(* Logix 5000 project; controller CIP vendor 1 type 14 code 106 rev 20.12; software revision 20.06; part 10 of 13 *)
(* tags used below, declared in another part *)
   MOA_OFF : DINT[10];
   MOA_ON : DINT[10];
   PV_Output_Status : INT[10];
   PV_Output_Status_IND : INT[10,16];
   PV_Status_Bit : BOOL;
   PV_Valve_Input_Status_IND : INT[10,16];
(* MainProgram, continued *)

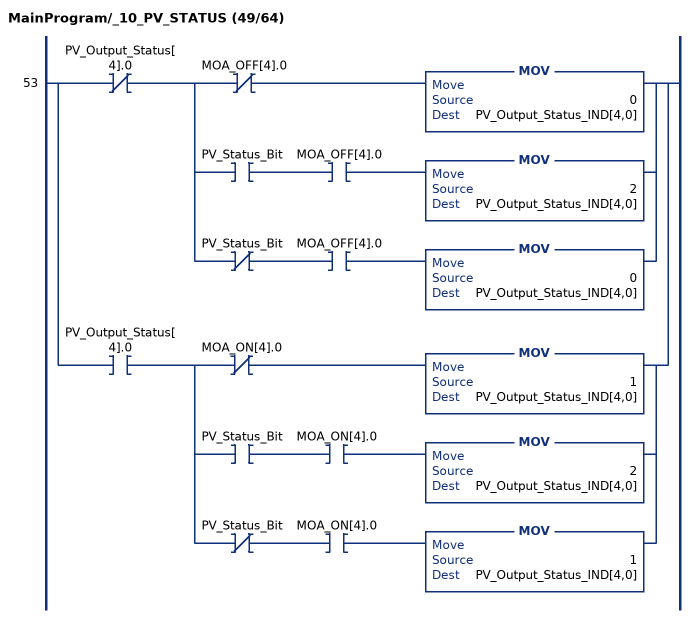
   [picture p181: MainProgram/_10_PV_STATUS rungs 53-53]
   53: [XIO(PV_Output_Status[4].0) [XIO(MOA_OFF[4].0) MOV(0,PV_Output_Status_IND[4,0]) ,XIC(PV_Status_Bit) XIC(MOA_OFF[4].0) MOV(2,PV_Output_Status_IND[4,0]) ,XIO(PV_Status_Bit) XIC(MOA_OFF[4].0) MOV(0,PV_Output_Status_IND[4,0]) ] ,XIC(PV_Output_Status[4].0) [XIO(MOA_ON[4].0) MOV(1,PV_Output_Status_IND[4,0]) ,XIC(PV_Status_Bit) XIC(MOA_ON[4].0) MOV(2,PV_Output_Status_IND[4,0]) ,XIO(PV_Status_Bit) XIC(MOA_ON[4].0) MOV(1,PV_Output_Status_IND[4,0]) ] ];
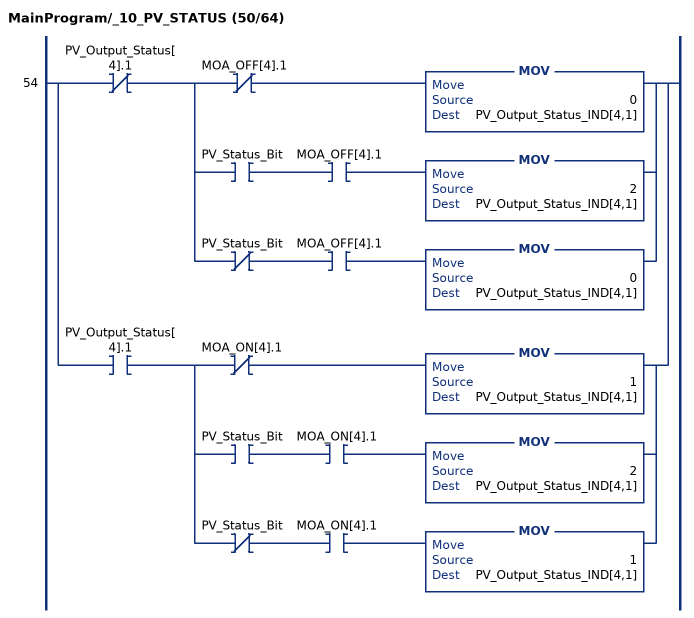
   54: [XIO(PV_Output_Status[4].1) [XIO(MOA_OFF[4].1) MOV(0,PV_Output_Status_IND[4,1]) ,XIC(PV_Status_Bit) XIC(MOA_OFF[4].1) MOV(2,PV_Output_Status_IND[4,1]) ,XIO(PV_Status_Bit) XIC(MOA_OFF[4].1) MOV(0,PV_Output_Status_IND[4,1]) ] ,XIC(PV_Output_Status[4].1) [XIO(MOA_ON[4].1) MOV(1,PV_Output_Status_IND[4,1]) ,XIC(PV_Status_Bit) XIC(MOA_ON[4].1) MOV(2,PV_Output_Status_IND[4,1]) ,XIO(PV_Status_Bit) XIC(MOA_ON[4].1) MOV(1,PV_Output_Status_IND[4,1]) ] ];
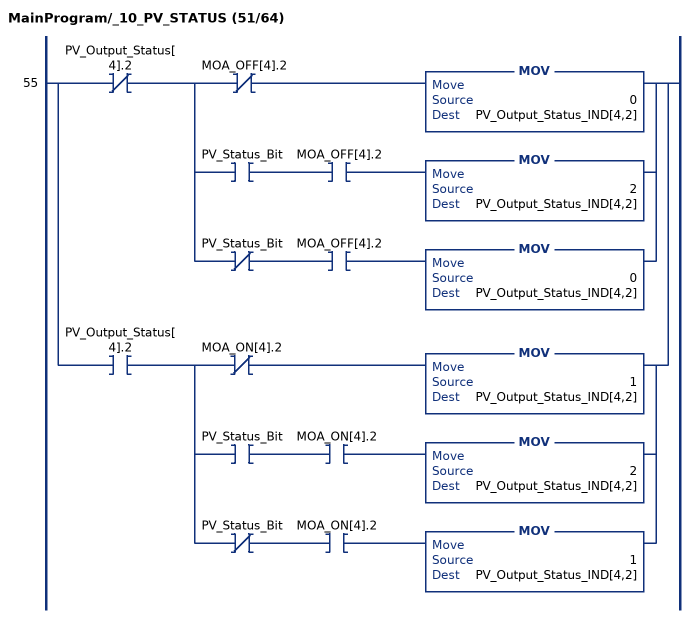
   55: [XIO(PV_Output_Status[4].2) [XIO(MOA_OFF[4].2) MOV(0,PV_Output_Status_IND[4,2]) ,XIC(PV_Status_Bit) XIC(MOA_OFF[4].2) MOV(2,PV_Output_Status_IND[4,2]) ,XIO(PV_Status_Bit) XIC(MOA_OFF[4].2) MOV(0,PV_Output_Status_IND[4,2]) ] ,XIC(PV_Output_Status[4].2) [XIO(MOA_ON[4].2) MOV(1,PV_Output_Status_IND[4,2]) ,XIC(PV_Status_Bit) XIC(MOA_ON[4].2) MOV(2,PV_Output_Status_IND[4,2]) ,XIO(PV_Status_Bit) XIC(MOA_ON[4].2) MOV(1,PV_Output_Status_IND[4,2]) ] ];
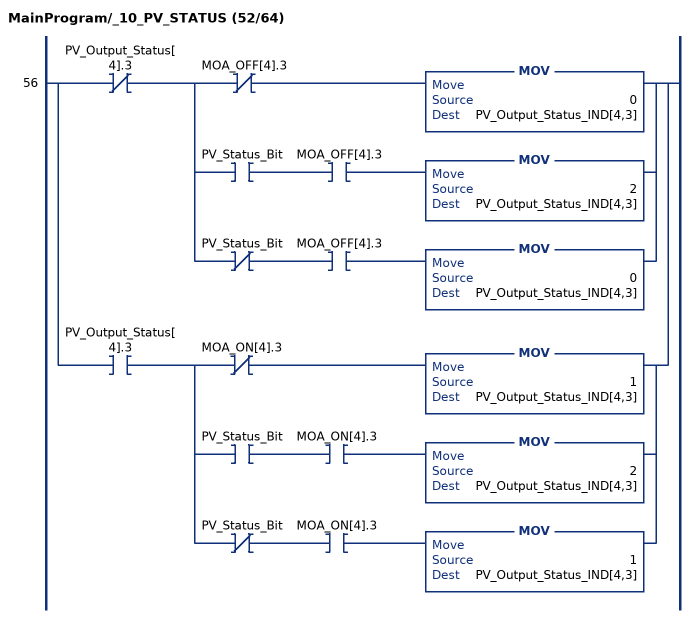
   56: [XIO(PV_Output_Status[4].3) [XIO(MOA_OFF[4].3) MOV(0,PV_Output_Status_IND[4,3]) ,XIC(PV_Status_Bit) XIC(MOA_OFF[4].3) MOV(2,PV_Output_Status_IND[4,3]) ,XIO(PV_Status_Bit) XIC(MOA_OFF[4].3) MOV(0,PV_Output_Status_IND[4,3]) ] ,XIC(PV_Output_Status[4].3) [XIO(MOA_ON[4].3) MOV(1,PV_Output_Status_IND[4,3]) ,XIC(PV_Status_Bit) XIC(MOA_ON[4].3) MOV(2,PV_Output_Status_IND[4,3]) ,XIO(PV_Status_Bit) XIC(MOA_ON[4].3) MOV(1,PV_Output_Status_IND[4,3]) ] ];
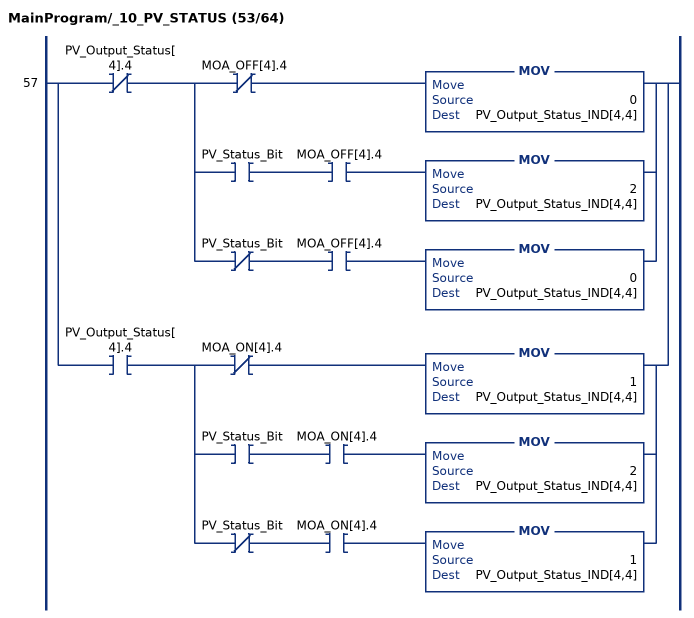
   57: [XIO(PV_Output_Status[4].4) [XIO(MOA_OFF[4].4) MOV(0,PV_Output_Status_IND[4,4]) ,XIC(PV_Status_Bit) XIC(MOA_OFF[4].4) MOV(2,PV_Output_Status_IND[4,4]) ,XIO(PV_Status_Bit) XIC(MOA_OFF[4].4) MOV(0,PV_Output_Status_IND[4,4]) ] ,XIC(PV_Output_Status[4].4) [XIO(MOA_ON[4].4) MOV(1,PV_Output_Status_IND[4,4]) ,XIC(PV_Status_Bit) XIC(MOA_ON[4].4) MOV(2,PV_Output_Status_IND[4,4]) ,XIO(PV_Status_Bit) XIC(MOA_ON[4].4) MOV(1,PV_Output_Status_IND[4,4]) ] ];
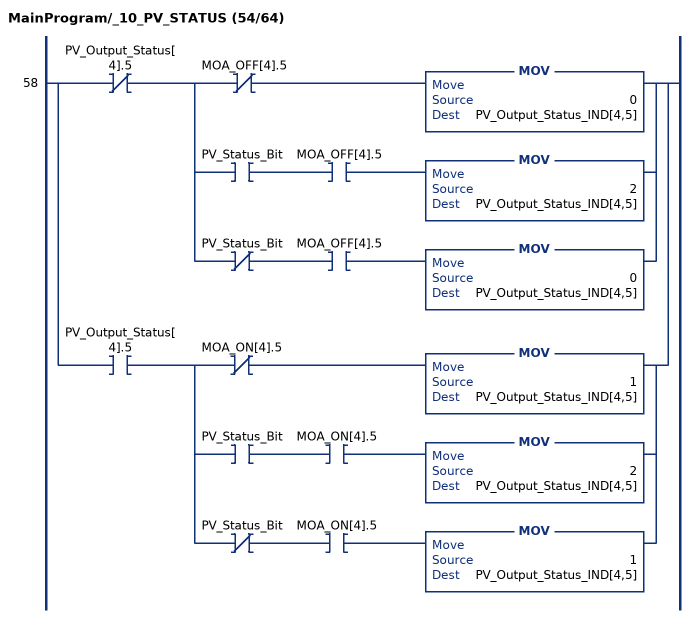
   58: [XIO(PV_Output_Status[4].5) [XIO(MOA_OFF[4].5) MOV(0,PV_Output_Status_IND[4,5]) ,XIC(PV_Status_Bit) XIC(MOA_OFF[4].5) MOV(2,PV_Output_Status_IND[4,5]) ,XIO(PV_Status_Bit) XIC(MOA_OFF[4].5) MOV(0,PV_Output_Status_IND[4,5]) ] ,XIC(PV_Output_Status[4].5) [XIO(MOA_ON[4].5) MOV(1,PV_Output_Status_IND[4,5]) ,XIC(PV_Status_Bit) XIC(MOA_ON[4].5) MOV(2,PV_Output_Status_IND[4,5]) ,XIO(PV_Status_Bit) XIC(MOA_ON[4].5) MOV(1,PV_Output_Status_IND[4,5]) ] ];
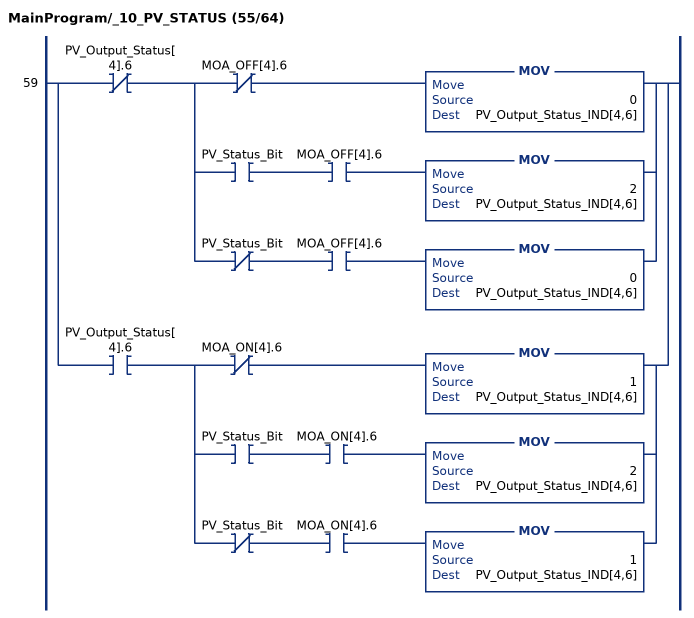
   59: [XIO(PV_Output_Status[4].6) [XIO(MOA_OFF[4].6) MOV(0,PV_Output_Status_IND[4,6]) ,XIC(PV_Status_Bit) XIC(MOA_OFF[4].6) MOV(2,PV_Output_Status_IND[4,6]) ,XIO(PV_Status_Bit) XIC(MOA_OFF[4].6) MOV(0,PV_Output_Status_IND[4,6]) ] ,XIC(PV_Output_Status[4].6) [XIO(MOA_ON[4].6) MOV(1,PV_Output_Status_IND[4,6]) ,XIC(PV_Status_Bit) XIC(MOA_ON[4].6) MOV(2,PV_Output_Status_IND[4,6]) ,XIO(PV_Status_Bit) XIC(MOA_ON[4].6) MOV(1,PV_Output_Status_IND[4,6]) ] ];
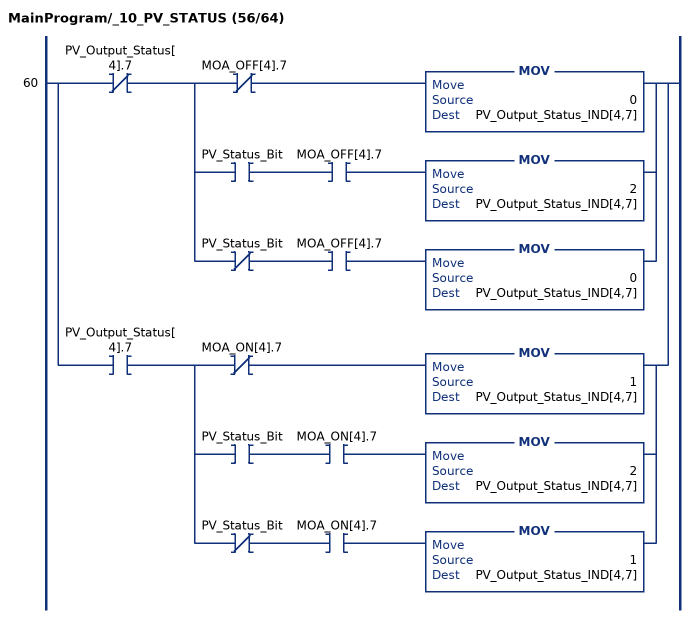
   60: [XIO(PV_Output_Status[4].7) [XIO(MOA_OFF[4].7) MOV(0,PV_Output_Status_IND[4,7]) ,XIC(PV_Status_Bit) XIC(MOA_OFF[4].7) MOV(2,PV_Output_Status_IND[4,7]) ,XIO(PV_Status_Bit) XIC(MOA_OFF[4].7) MOV(0,PV_Output_Status_IND[4,7]) ] ,XIC(PV_Output_Status[4].7) [XIO(MOA_ON[4].7) MOV(1,PV_Output_Status_IND[4,7]) ,XIC(PV_Status_Bit) XIC(MOA_ON[4].7) MOV(2,PV_Output_Status_IND[4,7]) ,XIO(PV_Status_Bit) XIC(MOA_ON[4].7) MOV(1,PV_Output_Status_IND[4,7]) ] ];
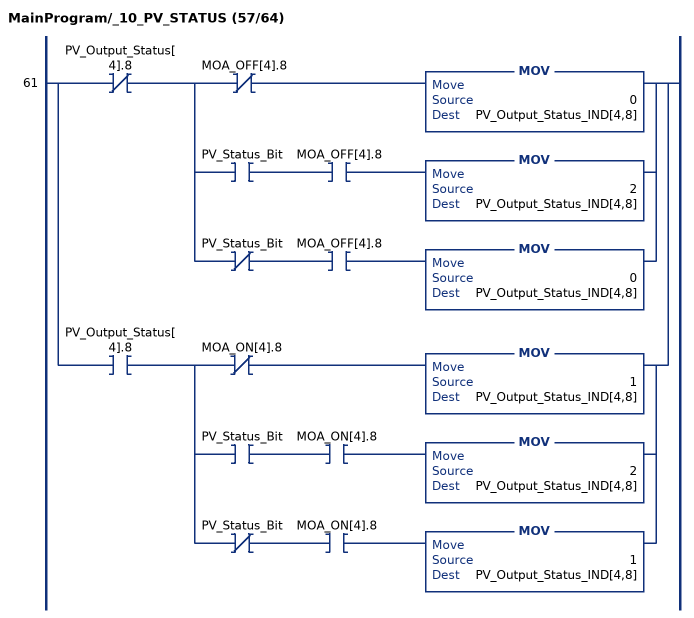
   61: [XIO(PV_Output_Status[4].8) [XIO(MOA_OFF[4].8) MOV(0,PV_Output_Status_IND[4,8]) ,XIC(PV_Status_Bit) XIC(MOA_OFF[4].8) MOV(2,PV_Output_Status_IND[4,8]) ,XIO(PV_Status_Bit) XIC(MOA_OFF[4].8) MOV(0,PV_Output_Status_IND[4,8]) ] ,XIC(PV_Output_Status[4].8) [XIO(MOA_ON[4].8) MOV(1,PV_Output_Status_IND[4,8]) ,XIC(PV_Status_Bit) XIC(MOA_ON[4].8) MOV(2,PV_Output_Status_IND[4,8]) ,XIO(PV_Status_Bit) XIC(MOA_ON[4].8) MOV(1,PV_Output_Status_IND[4,8]) ] ];
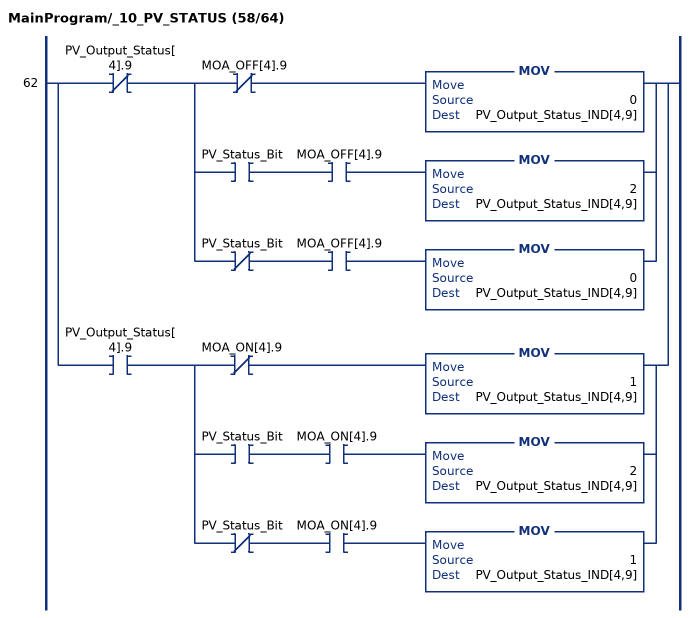
   62: [XIO(PV_Output_Status[4].9) [XIO(MOA_OFF[4].9) MOV(0,PV_Output_Status_IND[4,9]) ,XIC(PV_Status_Bit) XIC(MOA_OFF[4].9) MOV(2,PV_Output_Status_IND[4,9]) ,XIO(PV_Status_Bit) XIC(MOA_OFF[4].9) MOV(0,PV_Output_Status_IND[4,9]) ] ,XIC(PV_Output_Status[4].9) [XIO(MOA_ON[4].9) MOV(1,PV_Output_Status_IND[4,9]) ,XIC(PV_Status_Bit) XIC(MOA_ON[4].9) MOV(2,PV_Output_Status_IND[4,9]) ,XIO(PV_Status_Bit) XIC(MOA_ON[4].9) MOV(1,PV_Output_Status_IND[4,9]) ] ];
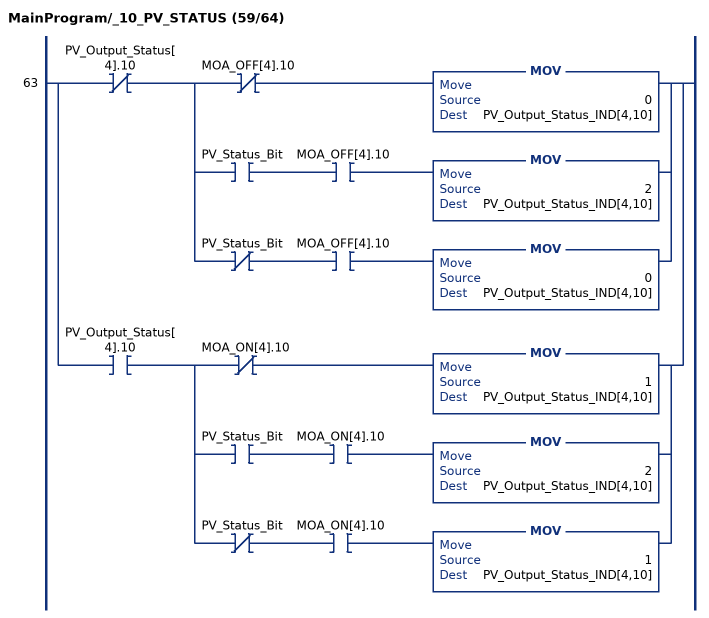
   63: [XIO(PV_Output_Status[4].10) [XIO(MOA_OFF[4].10) MOV(0,PV_Output_Status_IND[4,10]) ,XIC(PV_Status_Bit) XIC(MOA_OFF[4].10) MOV(2,PV_Output_Status_IND[4,10]) ,XIO(PV_Status_Bit) XIC(MOA_OFF[4].10) MOV(0,PV_Output_Status_IND[4,10]) ] ,XIC(PV_Output_Status[4].10) [XIO(MOA_ON[4].10) MOV(1,PV_Output_Status_IND[4,10]) ,XIC(PV_Status_Bit) XIC(MOA_ON[4].10) MOV(2,PV_Output_Status_IND[4,10]) ,XIO(PV_Status_Bit) XIC(MOA_ON[4].10) MOV(1,PV_Output_Status_IND[4,10]) ] ];
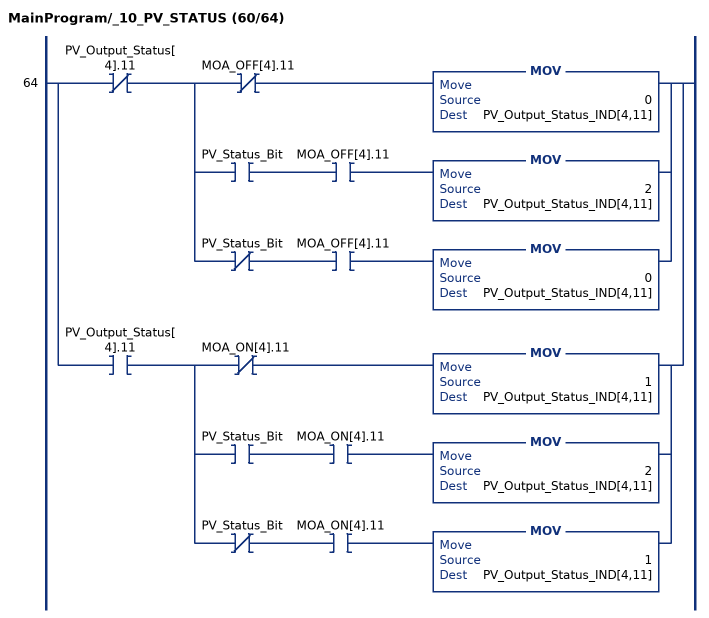
   64: [XIO(PV_Output_Status[4].11) [XIO(MOA_OFF[4].11) MOV(0,PV_Output_Status_IND[4,11]) ,XIC(PV_Status_Bit) XIC(MOA_OFF[4].11) MOV(2,PV_Output_Status_IND[4,11]) ,XIO(PV_Status_Bit) XIC(MOA_OFF[4].11) MOV(0,PV_Output_Status_IND[4,11]) ] ,XIC(PV_Output_Status[4].11) [XIO(MOA_ON[4].11) MOV(1,PV_Output_Status_IND[4,11]) ,XIC(PV_Status_Bit) XIC(MOA_ON[4].11) MOV(2,PV_Output_Status_IND[4,11]) ,XIO(PV_Status_Bit) XIC(MOA_ON[4].11) MOV(1,PV_Output_Status_IND[4,11]) ] ];
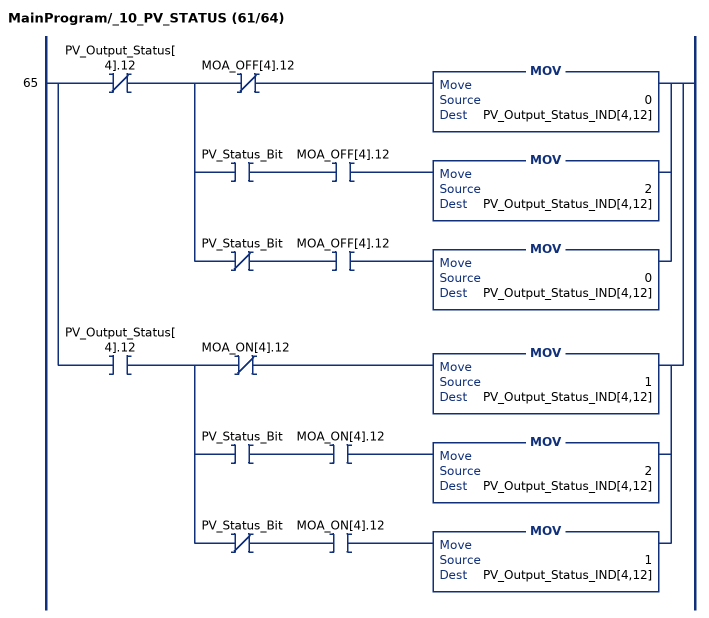
   65: [XIO(PV_Output_Status[4].12) [XIO(MOA_OFF[4].12) MOV(0,PV_Output_Status_IND[4,12]) ,XIC(PV_Status_Bit) XIC(MOA_OFF[4].12) MOV(2,PV_Output_Status_IND[4,12]) ,XIO(PV_Status_Bit) XIC(MOA_OFF[4].12) MOV(0,PV_Output_Status_IND[4,12]) ] ,XIC(PV_Output_Status[4].12) [XIO(MOA_ON[4].12) MOV(1,PV_Output_Status_IND[4,12]) ,XIC(PV_Status_Bit) XIC(MOA_ON[4].12) MOV(2,PV_Output_Status_IND[4,12]) ,XIO(PV_Status_Bit) XIC(MOA_ON[4].12) MOV(1,PV_Output_Status_IND[4,12]) ] ];
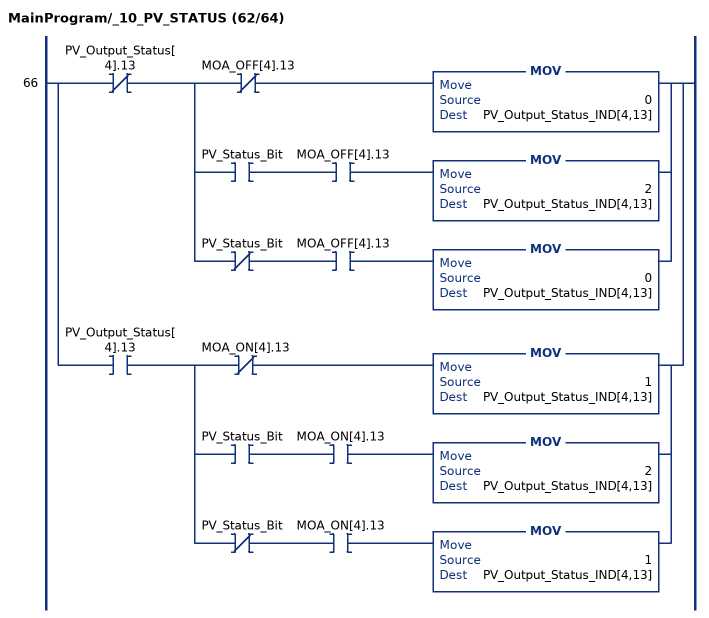
   66: [XIO(PV_Output_Status[4].13) [XIO(MOA_OFF[4].13) MOV(0,PV_Output_Status_IND[4,13]) ,XIC(PV_Status_Bit) XIC(MOA_OFF[4].13) MOV(2,PV_Output_Status_IND[4,13]) ,XIO(PV_Status_Bit) XIC(MOA_OFF[4].13) MOV(0,PV_Output_Status_IND[4,13]) ] ,XIC(PV_Output_Status[4].13) [XIO(MOA_ON[4].13) MOV(1,PV_Output_Status_IND[4,13]) ,XIC(PV_Status_Bit) XIC(MOA_ON[4].13) MOV(2,PV_Output_Status_IND[4,13]) ,XIO(PV_Status_Bit) XIC(MOA_ON[4].13) MOV(1,PV_Output_Status_IND[4,13]) ] ];
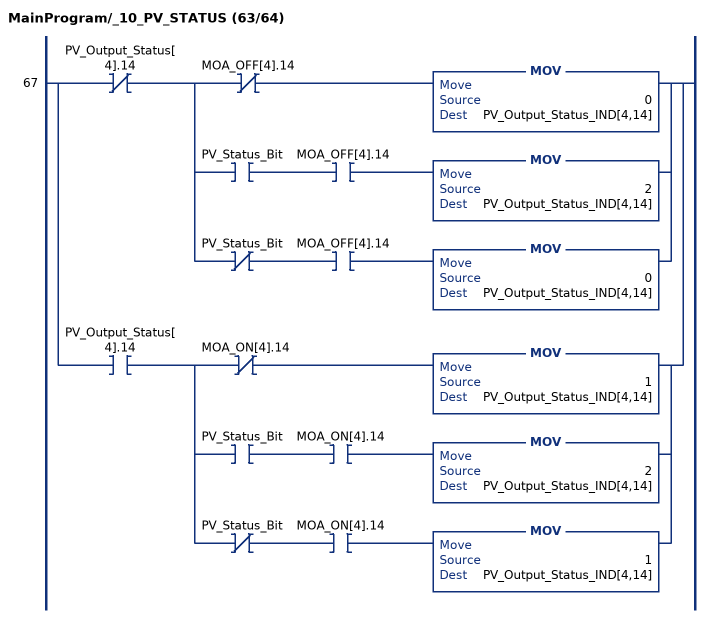
   67: [XIO(PV_Output_Status[4].14) [XIO(MOA_OFF[4].14) MOV(0,PV_Output_Status_IND[4,14]) ,XIC(PV_Status_Bit) XIC(MOA_OFF[4].14) MOV(2,PV_Output_Status_IND[4,14]) ,XIO(PV_Status_Bit) XIC(MOA_OFF[4].14) MOV(0,PV_Output_Status_IND[4,14]) ] ,XIC(PV_Output_Status[4].14) [XIO(MOA_ON[4].14) MOV(1,PV_Output_Status_IND[4,14]) ,XIC(PV_Status_Bit) XIC(MOA_ON[4].14) MOV(2,PV_Output_Status_IND[4,14]) ,XIO(PV_Status_Bit) XIC(MOA_ON[4].14) MOV(1,PV_Output_Status_IND[4,14]) ] ];
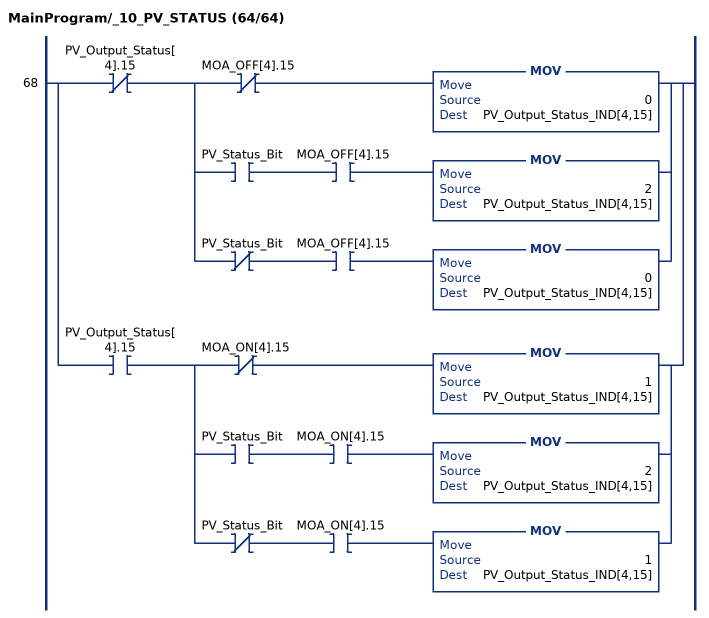
   68: [XIO(PV_Output_Status[4].15) [XIO(MOA_OFF[4].15) MOV(0,PV_Output_Status_IND[4,15]) ,XIC(PV_Status_Bit) XIC(MOA_OFF[4].15) MOV(2,PV_Output_Status_IND[4,15]) ,XIO(PV_Status_Bit) XIC(MOA_OFF[4].15) MOV(0,PV_Output_Status_IND[4,15]) ] ,XIC(PV_Output_Status[4].15) [XIO(MOA_ON[4].15) MOV(1,PV_Output_Status_IND[4,15]) ,XIC(PV_Status_Bit) XIC(MOA_ON[4].15) MOV(2,PV_Output_Status_IND[4,15]) ,XIO(PV_Status_Bit) XIC(MOA_ON[4].15) MOV(1,PV_Output_Status_IND[4,15]) ] ];
END_ROUTINE

ROUTINE _10_PV_VLV_STATUS   (* ladder *)
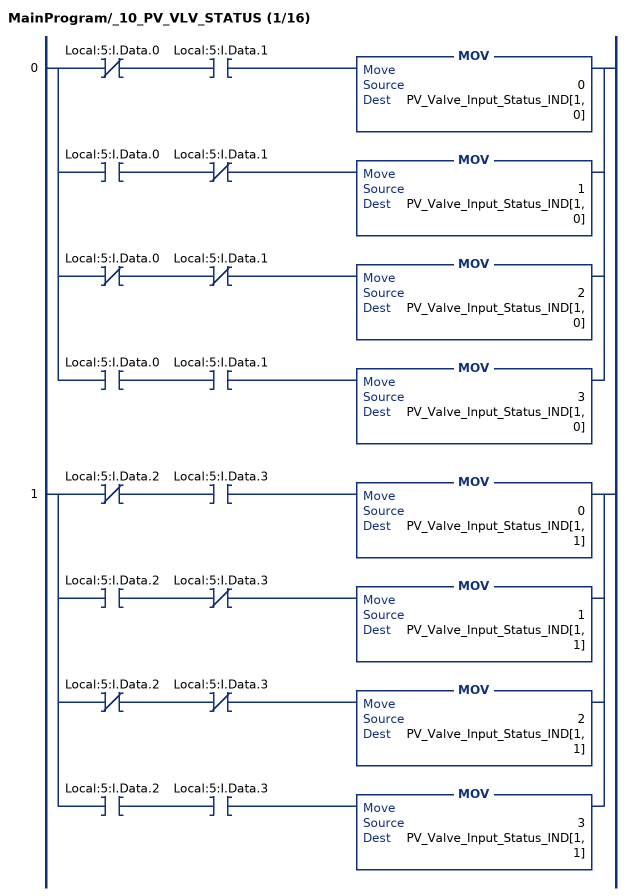
   0: [XIO(Local:5:I.Data.0) XIC(Local:5:I.Data.1) MOV(0,PV_Valve_Input_Status_IND[1,0]) ,XIC(Local:5:I.Data.0) XIO(Local:5:I.Data.1) MOV(1,PV_Valve_Input_Status_IND[1,0]) ,XIO(Local:5:I.Data.0) XIO(Local:5:I.Data.1) MOV(2,PV_Valve_Input_Status_IND[1,0]) ,XIC(Local:5:I.Data.0) XIC(Local:5:I.Data.1) MOV(3,PV_Valve_Input_Status_IND[1,0]) ];
   1: [XIO(Local:5:I.Data.2) XIC(Local:5:I.Data.3) MOV(0,PV_Valve_Input_Status_IND[1,1]) ,XIC(Local:5:I.Data.2) XIO(Local:5:I.Data.3) MOV(1,PV_Valve_Input_Status_IND[1,1]) ,XIO(Local:5:I.Data.2) XIO(Local:5:I.Data.3) MOV(2,PV_Valve_Input_Status_IND[1,1]) ,XIC(Local:5:I.Data.2) XIC(Local:5:I.Data.3) MOV(3,PV_Valve_Input_Status_IND[1,1]) ];
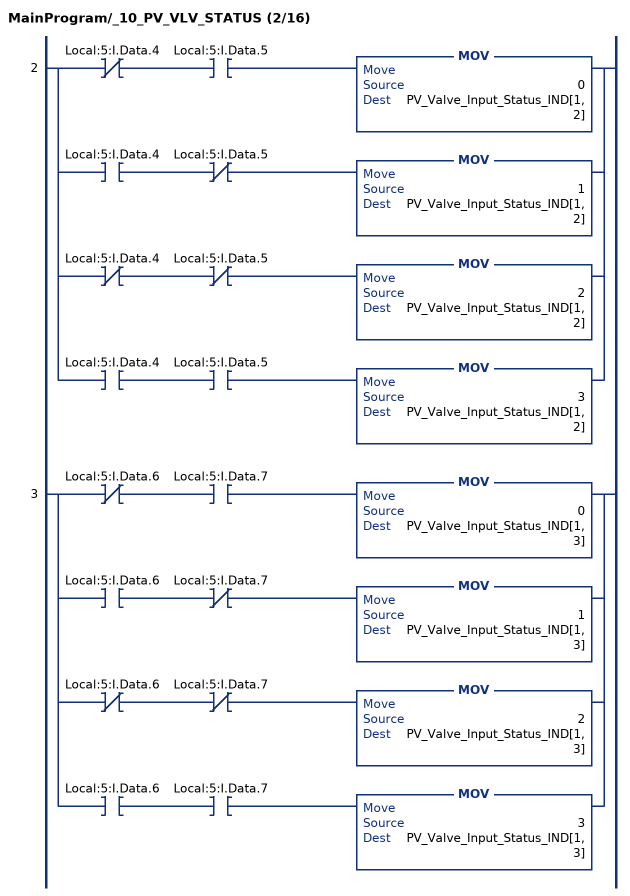
   2: [XIO(Local:5:I.Data.4) XIC(Local:5:I.Data.5) MOV(0,PV_Valve_Input_Status_IND[1,2]) ,XIC(Local:5:I.Data.4) XIO(Local:5:I.Data.5) MOV(1,PV_Valve_Input_Status_IND[1,2]) ,XIO(Local:5:I.Data.4) XIO(Local:5:I.Data.5) MOV(2,PV_Valve_Input_Status_IND[1,2]) ,XIC(Local:5:I.Data.4) XIC(Local:5:I.Data.5) MOV(3,PV_Valve_Input_Status_IND[1,2]) ];
   3: [XIO(Local:5:I.Data.6) XIC(Local:5:I.Data.7) MOV(0,PV_Valve_Input_Status_IND[1,3]) ,XIC(Local:5:I.Data.6) XIO(Local:5:I.Data.7) MOV(1,PV_Valve_Input_Status_IND[1,3]) ,XIO(Local:5:I.Data.6) XIO(Local:5:I.Data.7) MOV(2,PV_Valve_Input_Status_IND[1,3]) ,XIC(Local:5:I.Data.6) XIC(Local:5:I.Data.7) MOV(3,PV_Valve_Input_Status_IND[1,3]) ];
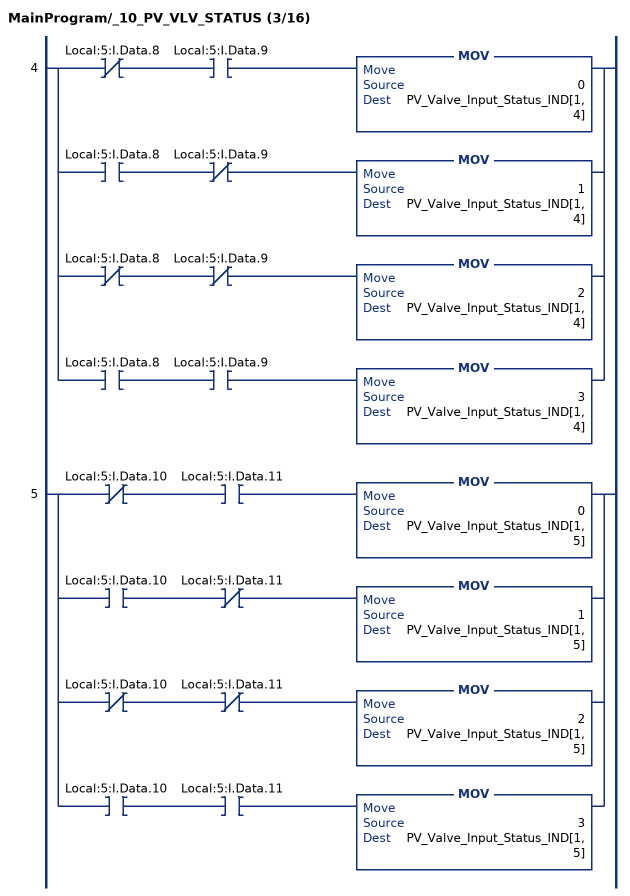
   4: [XIO(Local:5:I.Data.8) XIC(Local:5:I.Data.9) MOV(0,PV_Valve_Input_Status_IND[1,4]) ,XIC(Local:5:I.Data.8) XIO(Local:5:I.Data.9) MOV(1,PV_Valve_Input_Status_IND[1,4]) ,XIO(Local:5:I.Data.8) XIO(Local:5:I.Data.9) MOV(2,PV_Valve_Input_Status_IND[1,4]) ,XIC(Local:5:I.Data.8) XIC(Local:5:I.Data.9) MOV(3,PV_Valve_Input_Status_IND[1,4]) ];
   5: [XIO(Local:5:I.Data.10) XIC(Local:5:I.Data.11) MOV(0,PV_Valve_Input_Status_IND[1,5]) ,XIC(Local:5:I.Data.10) XIO(Local:5:I.Data.11) MOV(1,PV_Valve_Input_Status_IND[1,5]) ,XIO(Local:5:I.Data.10) XIO(Local:5:I.Data.11) MOV(2,PV_Valve_Input_Status_IND[1,5]) ,XIC(Local:5:I.Data.10) XIC(Local:5:I.Data.11) MOV(3,PV_Valve_Input_Status_IND[1,5]) ];
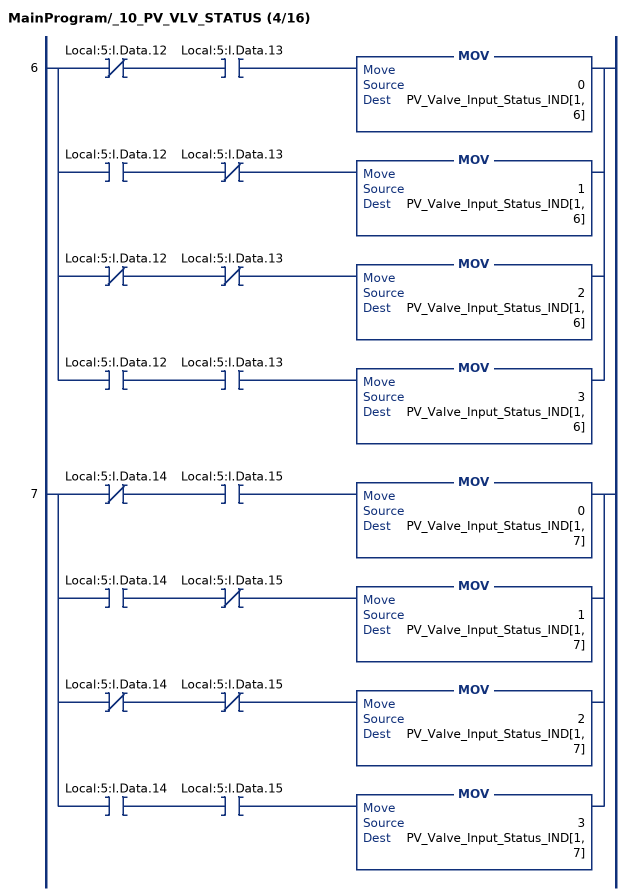
   6: [XIO(Local:5:I.Data.12) XIC(Local:5:I.Data.13) MOV(0,PV_Valve_Input_Status_IND[1,6]) ,XIC(Local:5:I.Data.12) XIO(Local:5:I.Data.13) MOV(1,PV_Valve_Input_Status_IND[1,6]) ,XIO(Local:5:I.Data.12) XIO(Local:5:I.Data.13) MOV(2,PV_Valve_Input_Status_IND[1,6]) ,XIC(Local:5:I.Data.12) XIC(Local:5:I.Data.13) MOV(3,PV_Valve_Input_Status_IND[1,6]) ];
   7: [XIO(Local:5:I.Data.14) XIC(Local:5:I.Data.15) MOV(0,PV_Valve_Input_Status_IND[1,7]) ,XIC(Local:5:I.Data.14) XIO(Local:5:I.Data.15) MOV(1,PV_Valve_Input_Status_IND[1,7]) ,XIO(Local:5:I.Data.14) XIO(Local:5:I.Data.15) MOV(2,PV_Valve_Input_Status_IND[1,7]) ,XIC(Local:5:I.Data.14) XIC(Local:5:I.Data.15) MOV(3,PV_Valve_Input_Status_IND[1,7]) ];
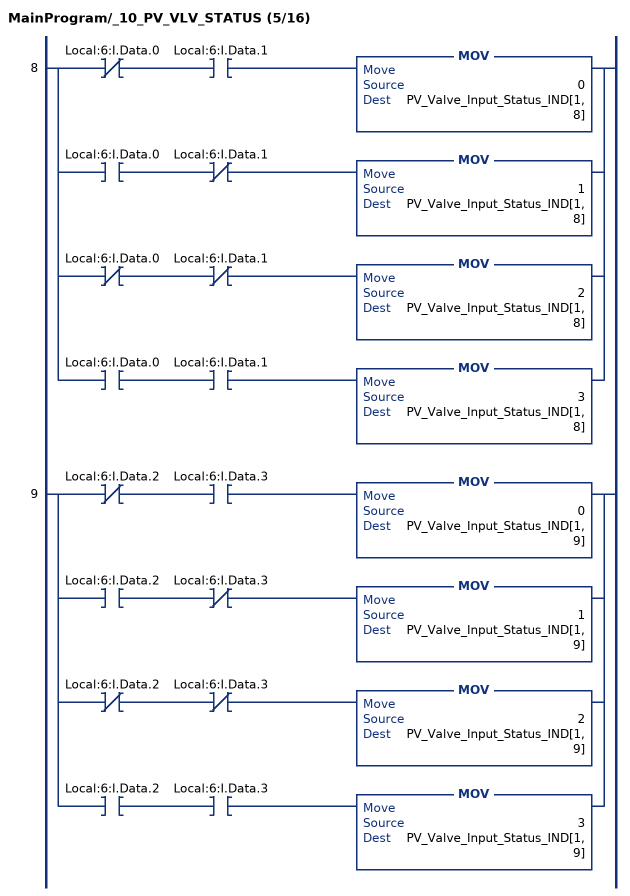
   8: [XIO(Local:6:I.Data.0) XIC(Local:6:I.Data.1) MOV(0,PV_Valve_Input_Status_IND[1,8]) ,XIC(Local:6:I.Data.0) XIO(Local:6:I.Data.1) MOV(1,PV_Valve_Input_Status_IND[1,8]) ,XIO(Local:6:I.Data.0) XIO(Local:6:I.Data.1) MOV(2,PV_Valve_Input_Status_IND[1,8]) ,XIC(Local:6:I.Data.0) XIC(Local:6:I.Data.1) MOV(3,PV_Valve_Input_Status_IND[1,8]) ];
   9: [XIO(Local:6:I.Data.2) XIC(Local:6:I.Data.3) MOV(0,PV_Valve_Input_Status_IND[1,9]) ,XIC(Local:6:I.Data.2) XIO(Local:6:I.Data.3) MOV(1,PV_Valve_Input_Status_IND[1,9]) ,XIO(Local:6:I.Data.2) XIO(Local:6:I.Data.3) MOV(2,PV_Valve_Input_Status_IND[1,9]) ,XIC(Local:6:I.Data.2) XIC(Local:6:I.Data.3) MOV(3,PV_Valve_Input_Status_IND[1,9]) ];
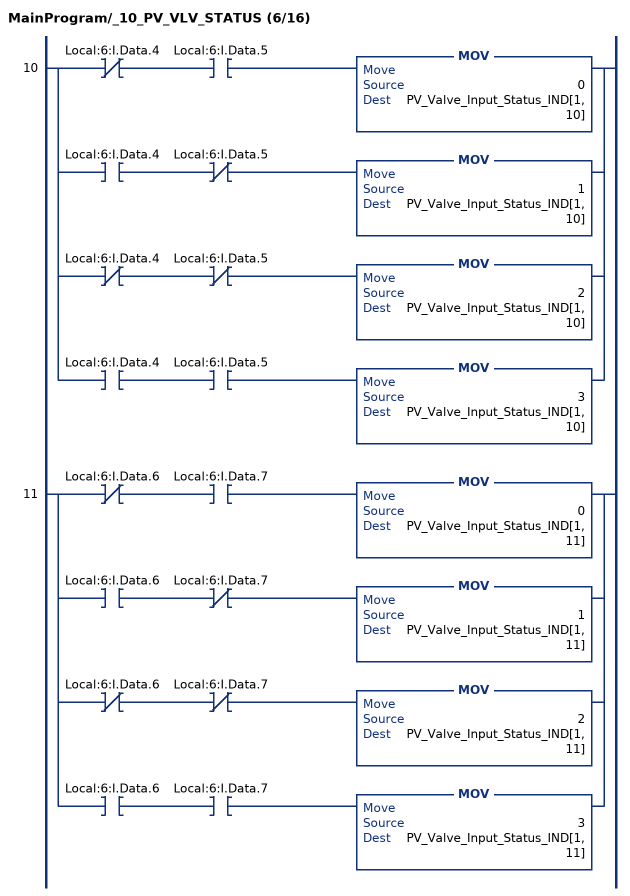
   10: [XIO(Local:6:I.Data.4) XIC(Local:6:I.Data.5) MOV(0,PV_Valve_Input_Status_IND[1,10]) ,XIC(Local:6:I.Data.4) XIO(Local:6:I.Data.5) MOV(1,PV_Valve_Input_Status_IND[1,10]) ,XIO(Local:6:I.Data.4) XIO(Local:6:I.Data.5) MOV(2,PV_Valve_Input_Status_IND[1,10]) ,XIC(Local:6:I.Data.4) XIC(Local:6:I.Data.5) MOV(3,PV_Valve_Input_Status_IND[1,10]) ];
   11: [XIO(Local:6:I.Data.6) XIC(Local:6:I.Data.7) MOV(0,PV_Valve_Input_Status_IND[1,11]) ,XIC(Local:6:I.Data.6) XIO(Local:6:I.Data.7) MOV(1,PV_Valve_Input_Status_IND[1,11]) ,XIO(Local:6:I.Data.6) XIO(Local:6:I.Data.7) MOV(2,PV_Valve_Input_Status_IND[1,11]) ,XIC(Local:6:I.Data.6) XIC(Local:6:I.Data.7) MOV(3,PV_Valve_Input_Status_IND[1,11]) ];
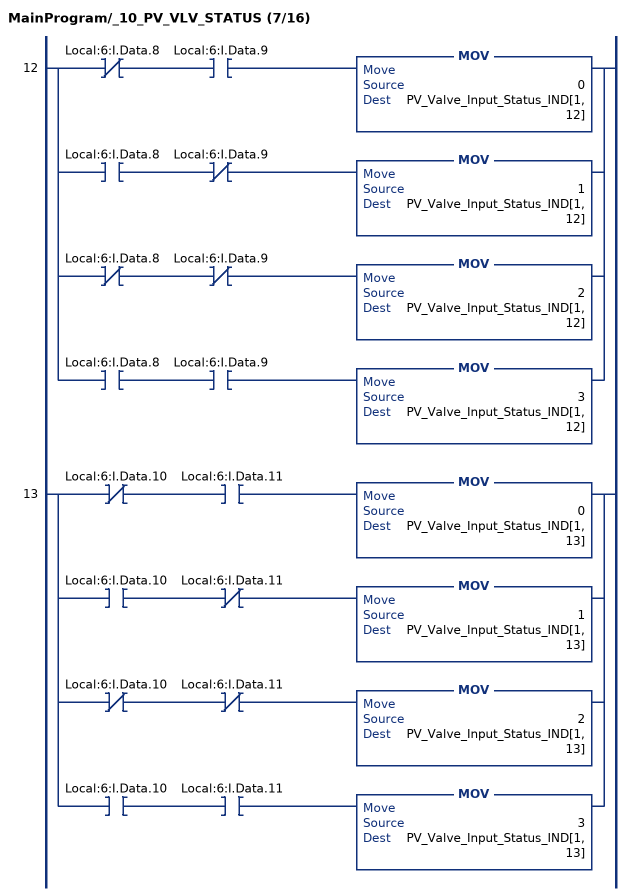
   12: [XIO(Local:6:I.Data.8) XIC(Local:6:I.Data.9) MOV(0,PV_Valve_Input_Status_IND[1,12]) ,XIC(Local:6:I.Data.8) XIO(Local:6:I.Data.9) MOV(1,PV_Valve_Input_Status_IND[1,12]) ,XIO(Local:6:I.Data.8) XIO(Local:6:I.Data.9) MOV(2,PV_Valve_Input_Status_IND[1,12]) ,XIC(Local:6:I.Data.8) XIC(Local:6:I.Data.9) MOV(3,PV_Valve_Input_Status_IND[1,12]) ];
   13: [XIO(Local:6:I.Data.10) XIC(Local:6:I.Data.11) MOV(0,PV_Valve_Input_Status_IND[1,13]) ,XIC(Local:6:I.Data.10) XIO(Local:6:I.Data.11) MOV(1,PV_Valve_Input_Status_IND[1,13]) ,XIO(Local:6:I.Data.10) XIO(Local:6:I.Data.11) MOV(2,PV_Valve_Input_Status_IND[1,13]) ,XIC(Local:6:I.Data.10) XIC(Local:6:I.Data.11) MOV(3,PV_Valve_Input_Status_IND[1,13]) ];
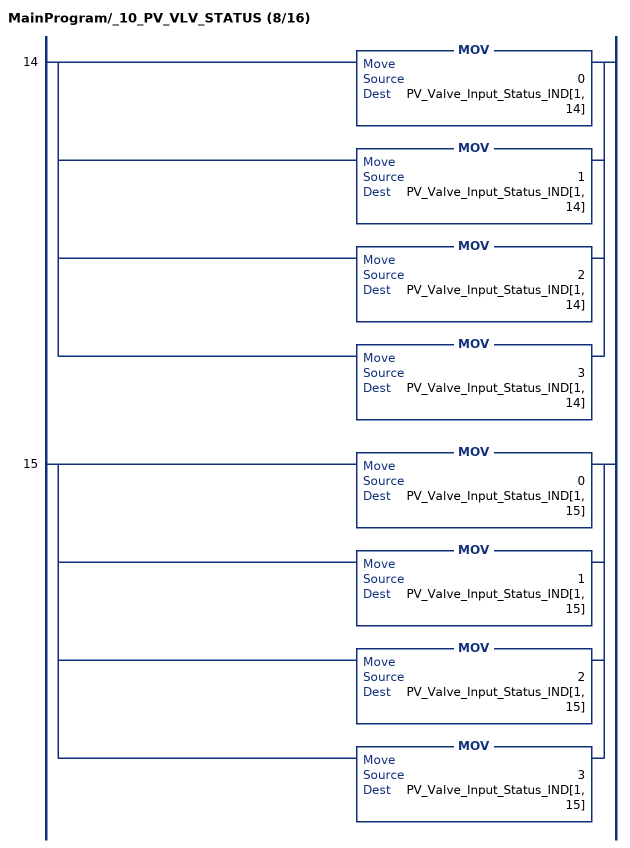
   14: [MOV(0,PV_Valve_Input_Status_IND[1,14]) ,MOV(1,PV_Valve_Input_Status_IND[1,14]) ,MOV(2,PV_Valve_Input_Status_IND[1,14]) ,MOV(3,PV_Valve_Input_Status_IND[1,14]) ];
   15: [MOV(0,PV_Valve_Input_Status_IND[1,15]) ,MOV(1,PV_Valve_Input_Status_IND[1,15]) ,MOV(2,PV_Valve_Input_Status_IND[1,15]) ,MOV(3,PV_Valve_Input_Status_IND[1,15]) ];
